(* IEC 61131-3 sources: codesys-ai-industrial-robot-control/plc/src/Equipment, 8 files *)

(* ---- FB_Bin.st ---- *)
(*
    FB_Bin
    Purpose : Output bin: counts placed parts and reports the full sensor.
    Inputs  : eBin - which bin; xFullSensor; xPlaced - rising edge = one part placed
    Outputs : uiCount, xFull
    Methods : Empty() - operator emptied the bin
*)
FUNCTION_BLOCK FB_Bin
VAR_INPUT
    eBin : E_Bin;
    xFullSensor : BOOL;
    xPlaced : BOOL;
END_VAR
VAR_OUTPUT
    uiCount : UINT;
    xFull : BOOL;
END_VAR
VAR
    rtPlaced : R_TRIG;
END_VAR

rtPlaced(CLK := xPlaced);
IF rtPlaced.Q THEN
    uiCount := uiCount + 1;
END_IF
xFull := xFullSensor;

(* ---- FB_CameraTrigger.st ---- *)
(*
    FB_CameraTrigger
    Purpose : On the PE1 photo-eye edge, assigns a new part id and publishes a capture request
              (with the conveyor position) for the vision service.
    Outputs : stCapture (udiSeq increments per request), xNewPart (one cycle), udiNewPartId
*)
FUNCTION_BLOCK FB_CameraTrigger
VAR_INPUT
    xPE1Rising : BOOL;
    lrBeltPos : LREAL;
END_VAR
VAR_OUTPUT
    stCapture : ST_CaptureMsg;
    xNewPart : BOOL;
    udiNewPartId : UDINT;
END_VAR

xNewPart := xPE1Rising;
IF xPE1Rising THEN
    udiNewPartId := udiNewPartId + 1;
    stCapture.udiSeq := stCapture.udiSeq + 1;
    stCapture.udiPartId := udiNewPartId;
    stCapture.lrBeltPos := lrBeltPos;
END_IF

(* ---- FB_Conveyor.st ---- *)
(*
    FB_Conveyor
    Purpose : Conveyor belt on a SoftMotion axis: power, run at a velocity, halt, read back.
    In/Out  : Axis - the conveyor axis (Axis_Conveyor)
    Inputs  : xEnable - power; lrVelocity - belt speed [mm/s]; xRun - move (FALSE = halt)
    Outputs : xPowered, xAtSpeed, lrPosition [mm], lrActVelocity [mm/s]
    Alarms  : ConveyorError
*)
FUNCTION_BLOCK FB_Conveyor IMPLEMENTS I_Equipment
VAR_IN_OUT
    Axis : AXIS_REF_SM3;
END_VAR
VAR_INPUT
    xEnable : BOOL;
    lrVelocity : LREAL;
    xRun : BOOL;
    itfAlarms : I_AlarmSink;
END_VAR
VAR_OUTPUT
    xPowered : BOOL;
    xAtSpeed : BOOL;
    lrPosition : LREAL;
    lrActVelocity : LREAL;
END_VAR
VAR
    fbPower : MC_Power;
    fbMove : MC_MoveVelocity;
    fbHalt : MC_Halt;
    fbReset : MC_Reset;
    fbReadPos : MC_ReadActualPosition;
    fbReadVel : MC_ReadActualVelocity;
    lrLastVelocity : LREAL;
    xRestart : BOOL;
    xResetRequest : BOOL;
    eError : E_AlarmId;
END_VAR
VAR CONSTANT
    ACCELERATION : LREAL := 1000;      // [mm/s2]
    JERK : LREAL := 10000;             // [mm/s3]
END_VAR

fbPower(Axis := Axis, Enable := xEnable, bRegulatorOn := xEnable, bDriveStart := xEnable);
xPowered := fbPower.Status;

// A changed velocity needs a new rising edge on Execute: drop it for one cycle.
xRestart := xRun AND lrVelocity <> lrLastVelocity;
lrLastVelocity := lrVelocity;
fbMove(Axis := Axis,
       Execute := xRun AND xPowered AND NOT xRestart AND eError = E_AlarmId.None,
       Velocity := ABS(lrVelocity),
       Acceleration := ACCELERATION,
       Deceleration := ACCELERATION,
       Jerk := JERK,
       Direction := MC_Direction.positive);
fbHalt(Axis := Axis, Execute := NOT xRun AND xPowered, Deceleration := ACCELERATION, Jerk := JERK);
xAtSpeed := fbMove.InVelocity;

fbReadPos(Axis := Axis, Enable := TRUE);
fbReadVel(Axis := Axis, Enable := TRUE);
lrPosition := fbReadPos.Position;
lrActVelocity := fbReadVel.Velocity;

IF (fbPower.Error OR fbMove.Error OR fbHalt.Error) AND eError = E_AlarmId.None THEN
    eError := E_AlarmId.ConveyorError;
    IF itfAlarms <> 0 THEN
        itfAlarms.Raise(eError);
    END_IF
END_IF

fbReset(Axis := Axis, Execute := xResetRequest);
IF xResetRequest AND (fbReset.Done OR fbReset.Error) THEN
    xResetRequest := FALSE;
    IF fbReset.Done THEN
        IF itfAlarms <> 0 AND eError <> E_AlarmId.None THEN
            itfAlarms.Clear(eError);
        END_IF
        eError := E_AlarmId.None;
    END_IF
END_IF

(* ---- FB_JointMonitor.st ---- *)
(*
    FB_JointMonitor
    Purpose : Supervises the robot joints against the feedback of the digital twin's servo
              motors: following error per joint and freshness of the feedback.
    Inputs  : aSetpoint / aFeedback [deg], aTorque [Nm], udiFeedbackSeq (changes with every new
              feedback sample), udiSetpointSeq (number of the current setpoint sample, +1 per
              cycle), udiFeedbackForSeq (setpoint sample the feedback answers), xLoopback
              (feedback := setpoint, no staleness check), xActive (supervision on), itfAlarms
    Outputs : aFollowingError [deg], iWorstJoint (1..6, 0 = none), xWarn, xFault, xStale
    Latency : the feedback travels through OPC UA and the twin (tens of ms). The last
              HISTORY_SIZE setpoints are kept, and the feedback is compared with the setpoint it
              answers, so transport delay does not count as following error. A feedback older
              than the history (a bridge hiccup) cannot be judged and counts as no error; if the
              feedback stays that old for tFeedbackTimeout it is stale.
    Debounce: a following error counts after CONFIRM_CYCLES cycles in a row. OPC UA does not
              hand a write to the task atomically: for one cycle the new positions may meet the
              old sequence number (a torn sample), which must not abort the cell.
    Limits  : GVL_Params.lrFollowErrWarn / lrFollowErrFault / tFeedbackTimeout
    Alarms  : FollowingErrorWarn, FollowingErrorFault, FeedbackStale
*)
FUNCTION_BLOCK FB_JointMonitor
VAR_INPUT
    aSetpoint : ARRAY[1..6] OF LREAL;
    aFeedback : ARRAY[1..6] OF LREAL;
    aTorque : ARRAY[1..6] OF LREAL;
    udiFeedbackSeq : UDINT;
    udiSetpointSeq : UDINT;
    udiFeedbackForSeq : UDINT;
    xLoopback : BOOL;
    xActive : BOOL;
    itfAlarms : I_AlarmSink;
END_VAR
VAR_OUTPUT
    aFollowingError : ARRAY[1..6] OF LREAL;
    iWorstJoint : INT;
    xWarn : BOOL;
    xFault : BOOL;
    xStale : BOOL;
END_VAR
VAR
    i : INT;
    lrWorst : LREAL;
    udiLastSeq : UDINT;
    tonStale : TON;
    aHistory : ARRAY[0..HISTORY_SIZE - 1, 1..6] OF LREAL;
    udiSlot : UDINT;
    xFromHistory : BOOL;
    uiWarnCycles : UINT;
    uiFaultCycles : UINT;
END_VAR
VAR CONSTANT
    HISTORY_SIZE : UDINT := 128;            // setpoint samples kept (512 ms at 4 ms)
    CONFIRM_CYCLES : UINT := 3;             // following error must persist this long (12 ms)
END_VAR

udiSlot := udiSetpointSeq MOD HISTORY_SIZE;
FOR i := 1 TO 6 DO
    aHistory[udiSlot, i] := aSetpoint[i];
END_FOR
// UDINT arithmetic: a feedback that answers a future setpoint wraps to a large age.
xFromHistory := udiSetpointSeq - udiFeedbackForSeq < HISTORY_SIZE;
udiSlot := udiFeedbackForSeq MOD HISTORY_SIZE;

lrWorst := 0;
iWorstJoint := 0;
FOR i := 1 TO 6 DO
    IF xLoopback OR NOT xFromHistory THEN
        aFollowingError[i] := 0;           // nothing to compare with: no judgement
    ELSE
        aFollowingError[i] := ABS(aHistory[udiSlot, i] - aFeedback[i]);
    END_IF
    IF aFollowingError[i] > lrWorst THEN
        lrWorst := aFollowingError[i];
        iWorstJoint := i;
    END_IF
END_FOR

IF xActive AND lrWorst > GVL_Params.lrFollowErrWarn THEN
    uiWarnCycles := MIN(uiWarnCycles + 1, CONFIRM_CYCLES);
ELSE
    uiWarnCycles := 0;
END_IF
IF xActive AND lrWorst > GVL_Params.lrFollowErrFault THEN
    uiFaultCycles := MIN(uiFaultCycles + 1, CONFIRM_CYCLES);
ELSE
    uiFaultCycles := 0;
END_IF
xWarn := uiWarnCycles >= CONFIRM_CYCLES;
xFault := uiFaultCycles >= CONFIRM_CYCLES;

// Feedback must keep arriving, and answer a setpoint still in the history, while supervised.
tonStale(IN := xActive AND NOT xLoopback AND (udiFeedbackSeq = udiLastSeq OR NOT xFromHistory),
         PT := GVL_Params.tFeedbackTimeout);
udiLastSeq := udiFeedbackSeq;
xStale := tonStale.Q;
xFault := xFault OR xStale;

IF itfAlarms <> 0 THEN
    IF xWarn THEN itfAlarms.Raise(E_AlarmId.FollowingErrorWarn); ELSE itfAlarms.Clear(E_AlarmId.FollowingErrorWarn); END_IF
    IF xFault AND NOT xStale THEN itfAlarms.Raise(E_AlarmId.FollowingErrorFault); ELSE itfAlarms.Clear(E_AlarmId.FollowingErrorFault); END_IF
    IF xStale THEN itfAlarms.Raise(E_AlarmId.FeedbackStale); ELSE itfAlarms.Clear(E_AlarmId.FeedbackStale); END_IF
END_IF

(* ---- FB_PhotoEye.st ---- *)
(*
    FB_PhotoEye
    Purpose : Debounced photo-eye with a rising-edge pulse.
    Inputs  : xRaw - sensor signal (TRUE = beam blocked); tDebounce - on/off filter time
    Outputs : xBlocked - debounced state; xRising - TRUE for one cycle when it becomes blocked
*)
FUNCTION_BLOCK FB_PhotoEye
VAR_INPUT
    xRaw : BOOL;
    tDebounce : TIME := T#10MS;
END_VAR
VAR_OUTPUT
    xBlocked : BOOL;
    xRising : BOOL;
END_VAR
VAR
    tonOn : TON;
    tonOff : TON;
END_VAR

tonOn(IN := xRaw, PT := tDebounce);
tonOff(IN := NOT xRaw, PT := tDebounce);
xRising := FALSE;
IF tonOn.Q AND NOT xBlocked THEN
    xBlocked := TRUE;
    xRising := TRUE;
ELSIF tonOff.Q THEN
    xBlocked := FALSE;
END_IF

(* ---- FB_Robot.st ---- *)
(*
    FB_Robot
    Purpose : The 6-axis robot (SoftMotion axis group) behind a PLCopen-style command interface.
    In/Out  : AxisGroup - AxisGroup_Robot
    Inputs  : xEnable - power and enable the group
              eCmd + stTarget - command, started by a rising edge of xExecute
              lrOverride - speed override ]0, 1] for all movements
    Outputs : xReady (enabled, no error), xBusy / xDone / xError of the running command,
              eSmcError, xMoving, stActAcs, stActMcs, aSetAcs[1..6] (joint setpoints, deg)
    Alarms  : AxisGroupError
    Lag     : SoftMotion's own TCP lag check compares the virtual drives' actual position, which
              trails the setpoint by one task cycle by design; its default (1 mm) trips at speed
              with Windows task jitter. MAX_TCP_LAG covers that; the real following error of the
              servo motors is supervised by FB_JointMonitor against the twin's feedback.
    Reset   : MC_GroupReset answers "no error to reset" when the group already left ErrorStop;
              that is a successful reset (otherwise the fault, and Clearing, would never end).
              The group is enabled only while it is disabled: re-enabling a group that a reset
              left enabled is an error of MC_GroupEnable.
    Note    : call once per cycle in the SoftMotion bus cycle task.
*)
FUNCTION_BLOCK FB_Robot IMPLEMENTS I_Equipment
VAR_IN_OUT
    AxisGroup : AXIS_GROUP_REF_SM3;
END_VAR
VAR_INPUT
    xEnable : BOOL;
    eCmd : E_RobotCmd;
    stTarget : SMC_POS_REF;
    xExecute : BOOL;
    lrOverride : LREAL := 1.0;
    itfAlarms : I_AlarmSink;
END_VAR
VAR_OUTPUT
    xReady : BOOL;
    xBusy : BOOL;
    xDone : BOOL;
    xError : BOOL;
    eSmcError : SMC_ERROR;
    xMoving : BOOL;
    stActAcs : SMC_POS_REF;
    stActMcs : SMC_POS_REF;
    aSetAcs : ARRAY[1..6] OF LREAL;
END_VAR
VAR CONSTANT
    MIN_OVERRIDE : LREAL := 0.01;
    STOP_DECELERATION : LREAL := 5000;     // path deceleration of a controlled stop [mm/s2]
    STOP_JERK : LREAL := 100000;           // path jerk of a controlled stop [mm/s3]
    MAX_TCP_LAG : LREAL := 10;             // SoftMotion TCP lag tolerance [mm]
    MAX_ORIENTATION_LAG : LREAL := 2;      // [deg]
    MAX_AXIS_LAG : LREAL := 2;             // per joint [deg]
END_VAR
VAR
    fbPower : SMC_GroupPower;
    fbEnable : MC_GroupEnable;
    fbReset : MC_GroupReset;
    fbStop : MC_GroupStop := (Deceleration := STOP_DECELERATION, Jerk := STOP_JERK);
    fbOverride : MC_GroupSetOverride;
    fbPtp : MC_MoveDirectAbsolute := (CoordSystem := SMC_COORD_SYSTEM.ACS);
    fbLin : MC_MoveLinearAbsolute;
    fbReadAcs : MC_GroupReadActualPosition := (Enable := TRUE, CoordSystem := SMC_COORD_SYSTEM.ACS);
    fbReadMcs : MC_GroupReadActualPosition := (Enable := TRUE, CoordSystem := SMC_COORD_SYSTEM.MCS);
    fbReadSet : SMC_GroupReadSetPosition := (Enable := TRUE, CoordSystem := SMC_COORD_SYSTEM.ACS);
    fbStatus : MC_GroupReadStatus := (Enable := TRUE);
    fbPathTol : SMC_GroupSetPathTolerance := (MaxPositionLag := MAX_TCP_LAG,
                                              MaxOrientationLag := MAX_ORIENTATION_LAG);
    rtExecute : R_TRIG;
    eActive : E_RobotCmd;
    xResetRequest : BOOL;
    xFault : BOOL;
    lrOverrideLimited : LREAL;
    xEnabled : BOOL;                       // powered and enabled, not in error
END_VAR

rtExecute(CLK := xExecute);
IF rtExecute.Q THEN
    eActive := eCmd;
ELSIF NOT xExecute THEN
    eActive := E_RobotCmd.None;
END_IF
IF eActive = E_RobotCmd.Reset THEN
    xResetRequest := TRUE;
END_IF

fbStatus(AxisGroup := AxisGroup);
fbPower(AxisGroup := AxisGroup, Enable := xEnable, bRegulatorOn := xEnable, bDriveStart := xEnable);
fbEnable(AxisGroup := AxisGroup,
         Execute := fbPower.Status AND NOT xResetRequest
                    AND (fbStatus.GroupDisabled OR fbEnable.Busy OR fbEnable.Done));
xEnabled := fbPower.Status AND fbStatus.Valid AND NOT fbStatus.GroupDisabled
            AND NOT fbStatus.GroupErrorStop;
fbPathTol.MaxAxisLag.a0 := MAX_AXIS_LAG;
fbPathTol.MaxAxisLag.a1 := MAX_AXIS_LAG;
fbPathTol.MaxAxisLag.a2 := MAX_AXIS_LAG;
fbPathTol.MaxAxisLag.a3 := MAX_AXIS_LAG;
fbPathTol.MaxAxisLag.a4 := MAX_AXIS_LAG;
fbPathTol.MaxAxisLag.a5 := MAX_AXIS_LAG;
fbPathTol(AxisGroup := AxisGroup, Execute := xEnabled);   // again after every enable

lrOverrideLimited := LIMIT(MIN_OVERRIDE, lrOverride, 1.0);
fbOverride(AxisGroup := AxisGroup,
           Enable := xEnabled AND NOT fbStatus.GroupStopping,
           VelFactor := lrOverrideLimited,
           PathVelFactor := lrOverrideLimited);

fbPtp.Position := stTarget;
fbPtp.VelFactor := GVL_Params.lrPtpVelFactor;
IF eActive = E_RobotCmd.MovePtpMcs THEN
    fbPtp.CoordSystem := SMC_COORD_SYSTEM.MCS;
ELSE
    fbPtp.CoordSystem := SMC_COORD_SYSTEM.ACS;
END_IF
fbPtp(AxisGroup := AxisGroup, Execute := eActive = E_RobotCmd.MovePtpAcs OR eActive = E_RobotCmd.MovePtpMcs);

fbLin.Position := stTarget;
fbLin.Velocity := GVL_Params.lrLinVelocity;
fbLin.Acceleration := GVL_Params.lrLinAccel;
fbLin.Deceleration := GVL_Params.lrLinAccel;
fbLin.Jerk := GVL_Params.lrLinJerk;
IF eActive = E_RobotCmd.MoveLinPcs1 THEN
    fbLin.CoordSystem := SMC_COORD_SYSTEM.PCS_1;
ELSE
    fbLin.CoordSystem := SMC_COORD_SYSTEM.MCS;
END_IF
fbLin(AxisGroup := AxisGroup, Execute := eActive = E_RobotCmd.MoveLinMcs OR eActive = E_RobotCmd.MoveLinPcs1);

fbStop(AxisGroup := AxisGroup, Execute := eActive = E_RobotCmd.Stop);
fbReset(AxisGroup := AxisGroup, Execute := xResetRequest);
IF xResetRequest AND (fbReset.Done OR fbReset.Error) THEN
    xResetRequest := FALSE;
    IF fbReset.Done OR NOT fbStatus.GroupErrorStop THEN
        IF xFault AND itfAlarms <> 0 THEN
            itfAlarms.Clear(E_AlarmId.AxisGroupError);
        END_IF
        xFault := FALSE;
        eSmcError := SMC_ERROR.SMC_NO_ERROR;
    END_IF
    fbStatus(AxisGroup := AxisGroup);   // the fault check below must see the state after the reset
END_IF

fbReadAcs(AxisGroup := AxisGroup);
fbReadMcs(AxisGroup := AxisGroup);
fbReadSet(AxisGroup := AxisGroup);
stActAcs := fbReadAcs.Position;
stActMcs := fbReadMcs.Position;
aSetAcs[1] := fbReadSet.Position.a.a0;
aSetAcs[2] := fbReadSet.Position.a.a1;
aSetAcs[3] := fbReadSet.Position.a.a2;
aSetAcs[4] := fbReadSet.Position.a.a3;
aSetAcs[5] := fbReadSet.Position.a.a4;
aSetAcs[6] := fbReadSet.Position.a.a5;

CASE eActive OF
    E_RobotCmd.MovePtpAcs, E_RobotCmd.MovePtpMcs:
        xBusy := fbPtp.Busy; xDone := fbPtp.Done; xError := fbPtp.Error;
        IF fbPtp.Error THEN eSmcError := fbPtp.ErrorID; END_IF
    E_RobotCmd.MoveLinMcs, E_RobotCmd.MoveLinPcs1:
        xBusy := fbLin.Busy; xDone := fbLin.Done; xError := fbLin.Error;
        IF fbLin.Error THEN eSmcError := fbLin.ErrorID; END_IF
    E_RobotCmd.Stop:
        xBusy := fbStop.Busy; xDone := fbStop.Done; xError := fbStop.Error;
        IF fbStop.Error THEN eSmcError := fbStop.ErrorID; END_IF
    E_RobotCmd.Reset:
        xBusy := xResetRequest; xDone := NOT xResetRequest AND NOT xFault;
        xError := fbReset.Error AND fbStatus.GroupErrorStop;
ELSE
    xBusy := FALSE; xDone := FALSE; xError := FALSE;
END_CASE

IF (fbPower.Error OR fbEnable.Error OR fbStatus.GroupErrorStop OR xError) AND NOT xFault
   AND NOT xResetRequest THEN
    xFault := TRUE;
    IF eSmcError = SMC_ERROR.SMC_NO_ERROR THEN
        IF fbEnable.Error THEN eSmcError := fbEnable.ErrorID; ELSE eSmcError := fbPower.ErrorID; END_IF
    END_IF
    IF itfAlarms <> 0 THEN
        itfAlarms.Raise(E_AlarmId.AxisGroupError);
    END_IF
END_IF

xMoving := fbStatus.GroupMoving OR fbStatus.GroupStopping;
xReady := xEnabled AND NOT xFault;

(* ---- FB_SafetyMonitor.st ---- *)
(*
    FB_SafetyMonitor
    Purpose : Modelled safety logic (not certified): E-stop latch and safety door per mode.
    Inputs  : xEStopOk (TRUE = not pressed), xDoorClosed, eMode, xResetCmd, itfAlarms
    Outputs : xSafeToMove - motion allowed; xReducedSpeed - only reduced speed allowed
    Rules   : E-stop latches until xEStopOk AND xResetCmd. Door open in Production or
              Maintenance -> not safe (DoorOpen). Door open in Manual -> safe, reduced speed.
    Alarms  : EStop, DoorOpen
*)
FUNCTION_BLOCK FB_SafetyMonitor
VAR_INPUT
    xEStopOk : BOOL := TRUE;
    xDoorClosed : BOOL := TRUE;
    eMode : E_PackMLMode := E_PackMLMode.Production;
    xResetCmd : BOOL;
    itfAlarms : I_AlarmSink;
END_VAR
VAR_OUTPUT
    xSafeToMove : BOOL;
    xReducedSpeed : BOOL;
END_VAR
VAR
    xEStopLatched : BOOL;
    xDoorFault : BOOL;
END_VAR

IF NOT xEStopOk THEN
    xEStopLatched := TRUE;
ELSIF xResetCmd THEN
    xEStopLatched := FALSE;
END_IF

xDoorFault := NOT xDoorClosed AND eMode <> E_PackMLMode.Manual;
xSafeToMove := NOT xEStopLatched AND NOT xDoorFault;
xReducedSpeed := NOT xDoorClosed AND eMode = E_PackMLMode.Manual;

IF itfAlarms <> 0 THEN
    IF xEStopLatched THEN
        itfAlarms.Raise(E_AlarmId.EStop);
    ELSE
        itfAlarms.Clear(E_AlarmId.EStop);
    END_IF
    IF xDoorFault THEN
        itfAlarms.Raise(E_AlarmId.DoorOpen);
    ELSE
        itfAlarms.Clear(E_AlarmId.DoorOpen);
    END_IF
END_IF

(* ---- FB_VacuumGripper.st ---- *)
(*
    FB_VacuumGripper
    Purpose : Suction gripper: valve control with grip and loss supervision.
    Inputs  : xCmdVacuum, xVacuumOk (vacuum switch), tGripTimeout, itfAlarms
    Outputs : xValveOn, xHolding (vacuum on and OK)
    Errors  : VacuumNoGrip - commanded but not OK within tGripTimeout
              VacuumLost - was holding and lost vacuum while still commanded
*)
FUNCTION_BLOCK FB_VacuumGripper IMPLEMENTS I_Equipment
VAR_INPUT
    xCmdVacuum : BOOL;
    xVacuumOk : BOOL;
    tGripTimeout : TIME := T#500MS;
    itfAlarms : I_AlarmSink;
END_VAR
VAR_OUTPUT
    xValveOn : BOOL;
    xHolding : BOOL;
END_VAR
VAR
    tonGrip : TON;
    xWasHolding : BOOL;
    eError : E_AlarmId;
END_VAR

xValveOn := xCmdVacuum;
xHolding := xCmdVacuum AND xVacuumOk;

tonGrip(IN := xCmdVacuum AND NOT xVacuumOk AND NOT xWasHolding, PT := tGripTimeout);
IF tonGrip.Q AND eError = E_AlarmId.None THEN
    eError := E_AlarmId.VacuumNoGrip;
END_IF
IF xWasHolding AND xCmdVacuum AND NOT xVacuumOk AND eError = E_AlarmId.None THEN
    eError := E_AlarmId.VacuumLost;
END_IF

IF xHolding THEN
    xWasHolding := TRUE;
ELSIF NOT xCmdVacuum THEN
    xWasHolding := FALSE;
END_IF

IF eError <> E_AlarmId.None AND itfAlarms <> 0 THEN
    itfAlarms.Raise(eError);
END_IF
